Fanuc KAREL source: kt00026.KL

-- PROVISIONAL review KL for V770-1; original PC SHA256 247b8c3ce72dbd680a0f780a6a1b7390c90834b09a0120338ba43aaa4772aa64
-- Incomplete behavior may be omitted. Consult companion uncertainty JSON. Do not deploy.
PROGRAM KT00026
%NOLOCKGROUP
VAR
  I2 : INTEGER
  OUT : REAL
-- UNRESOLVED_DECL H1 type=002017
BEGIN
  -- UNRESOLVED_PC offsets 5-19; opcodes 2E,22,9D,33,B4
  -- UNRESOLVED_PC offsets 24-35; opcodes 2E,23
  -- UNRESOLVED_PC offsets 40-63; opcodes 22,9D,33,B3,21,52,64,23
  -- UNRESOLVED_PC offsets 68-72; opcodes 7F
END KT00026
